// TIA Portal project "Testing 1" (V18)

(* hardware
DEVICE "S7-1200 station_1"  S7-1200 Station
   slot 0: "Rack_0"  S7-1200 Rack  Rack  V1.0
   slot 1: "PLC_1"  CPU 1215C DC/DC/DC  6ES7 215-1AG40-0XB0  V4.6
   slot 2: "SM 1278_1"  4SI IO link  6ES7 278-4BD32-0XB0  V2.1
   slot 3: "DI 2/DQ 2x24VDC_1"  DI2/DQ2 signal board  6ES7 223-0BD30-0XB0  V1.0
*)

// ===== PLC "PLC_1"  CPU 1215C DC/DC/DC =====

VAR_GLOBAL   // PLC tag table "Default tag table"
   "err" AT %MW2 : Int;
END_VAR

VAR_GLOBAL   // PLC tag table "Tag table_1"
   "Marche" AT %M0.0 : Bool;
   "Web_CMD_StartMarche" AT %M0.1 : Bool;
   "Web_CMD_StopMarche" AT %M0.2 : Bool;
   "b1" AT %I1.3 : Bool;
   "b2" AT %I1.4 : Bool;
   "km1" AT %Q1.0 : Bool;
   "km2" AT %Q1.1 : Bool;
END_VAR

FUNCTION "test" : Void   // FC1, LAD
{ S7_Optimized_Access := 'TRUE' }
VERSION : 0.1
BEGIN

REGION Network 1
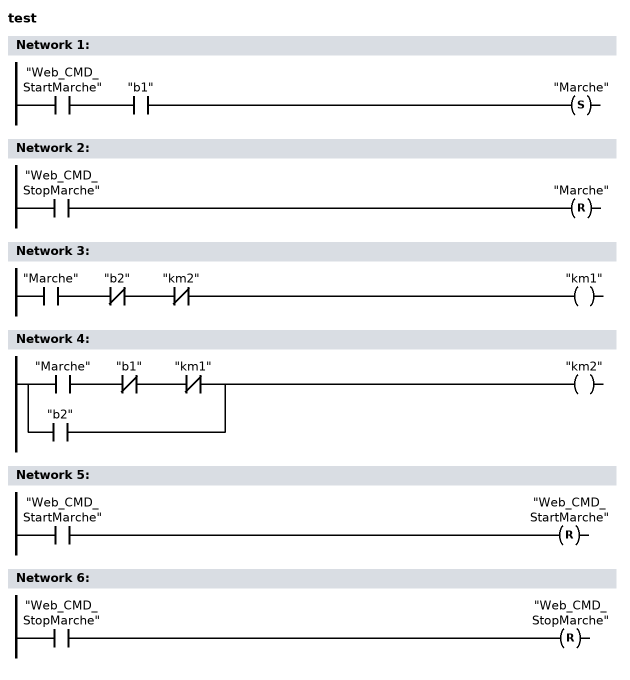
   RUNG wire#powerrail
      Contact( "Web_CMD_StartMarche" )
      Contact( "b1" )
      S_Coil( "Marche" )
   END_RUNG
   // the same network as SCL:
   IF "Web_CMD_StartMarche" AND "b1" THEN "Marche" := TRUE; END_IF;
END_REGION

REGION Network 2
   RUNG wire#powerrail
      Contact( "Web_CMD_StopMarche" )
      R_Coil( "Marche" )
   END_RUNG
   // the same network as SCL:
   IF "Web_CMD_StopMarche" THEN "Marche" := FALSE; END_IF;
END_REGION

REGION Network 3
   RUNG wire#powerrail
      Contact( "Marche" )
      I_Contact( "b2" )
      I_Contact( "km2" )
      Coil( "km1" )
   END_RUNG
   // the same network as SCL:
   "km1" := "Marche" AND NOT "b2" AND NOT "km2";
END_REGION

REGION Network 4
   RUNG wire#powerrail
      Contact( "Marche" )
      I_Contact( "b1" )
      I_Contact( "km1" )
      wire#w1
      Coil( "km2" )
   END_RUNG
   RUNG wire#powerrail
      Contact( "b2" )
   END_RUNG wire#w1
   // the same network as SCL:
   "km2" := ("Marche" AND NOT "b1" AND NOT "km1") OR "b2";
END_REGION

REGION Network 5
   RUNG wire#powerrail
      Contact( "Web_CMD_StartMarche" )
      R_Coil( "Web_CMD_StartMarche" )
   END_RUNG
   // the same network as SCL:
   IF "Web_CMD_StartMarche" THEN "Web_CMD_StartMarche" := FALSE; END_IF;
END_REGION

REGION Network 6
   RUNG wire#powerrail
      Contact( "Web_CMD_StopMarche" )
      R_Coil( "Web_CMD_StopMarche" )
   END_RUNG
   // the same network as SCL:
   IF "Web_CMD_StopMarche" THEN "Web_CMD_StopMarche" := FALSE; END_IF;
END_REGION
END_FUNCTION

ORGANIZATION_BLOCK "Main"   // OB1, LAD, ProgramCycle
TITLE = "Main Program Sweep (Cycle)"
{ S7_Optimized_Access := 'TRUE' }
VERSION : 0.1
   VAR_INPUT
      Initial_Call : Bool;   // Initial call of this OB
      Remanence : Bool;   // =True, if remanent data are available
   END_VAR
BEGIN

REGION Network 1
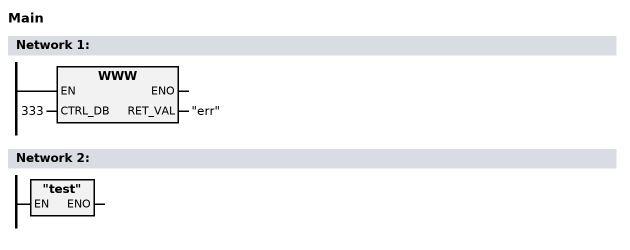
   "err" := WWW(CTRL_DB := 333);
END_REGION

REGION Network 2
   RUNG wire#powerrail
      "test"()
   END_RUNG
   // the same network as SCL:
   "test"();
END_REGION
END_ORGANIZATION_BLOCK